(* IEC 61131-3 sources: plc-iiot-stack/src/GVLs/Generated, 1 file *)

(* ---- GVL_IiotMap.gvl.st ---- *)
// AUTO-GENERATED by gen_plc_iiot.py — не редактировать; источник: schema/ (метрики, команды, тревоги)
// Назначение: размеры и таблицы настроек ПЛК-части IIoT-стека КНС-1: метрики телеметрии (топик
//             <site>/<area>/<unit>/<sPath>), белый список команд, тревоги перечня флагмана.
//             Индексы PT_<DEVICE>_<METRIC> — номера метрик в таблице POINT_CFG.
// Документ:   docs/plc_mqtt.md, раздел «Таблицы из схемы данных»
{attribute 'qualified_only'}
VAR_GLOBAL CONSTANT
    POINT_COUNT : DINT := 139;
    RULE_COUNT : DINT := 86;
    CMD_DEVICE_COUNT : DINT := 31;
    ALARM_COUNT : DINT := 88;
    ALARM_WORDS_COUNT : DINT := 28;

    // Метрики (schema/telemetry_catalog.csv)
    PT_P101_RUNNING : DINT := 1;
    PT_P101_STATE : DINT := 2;
    PT_P101_SPEED : DINT := 3;
    PT_P101_SPEED_REF : DINT := 4;
    PT_P101_RUN_HOURS : DINT := 5;
    PT_P101_STARTS : DINT := 6;
    PT_P101_STARTS_LAST_HOUR : DINT := 7;
    PT_P101_RUN_HOURS_MAINT : DINT := 8;
    PT_P101_STARTS_MAINT : DINT := 9;
    PT_P101_VFD_FAULT_CODE : DINT := 10;
    PT_P101_MODE : DINT := 11;
    PT_P101_NE107 : DINT := 12;
    PT_P102_RUNNING : DINT := 13;
    PT_P102_STATE : DINT := 14;
    PT_P102_SPEED : DINT := 15;
    PT_P102_SPEED_REF : DINT := 16;
    PT_P102_RUN_HOURS : DINT := 17;
    PT_P102_STARTS : DINT := 18;
    PT_P102_STARTS_LAST_HOUR : DINT := 19;
    PT_P102_RUN_HOURS_MAINT : DINT := 20;
    PT_P102_STARTS_MAINT : DINT := 21;
    PT_P102_VFD_FAULT_CODE : DINT := 22;
    PT_P102_MODE : DINT := 23;
    PT_P102_NE107 : DINT := 24;
    PT_P103_RUNNING : DINT := 25;
    PT_P103_STATE : DINT := 26;
    PT_P103_SPEED : DINT := 27;
    PT_P103_SPEED_REF : DINT := 28;
    PT_P103_RUN_HOURS : DINT := 29;
    PT_P103_STARTS : DINT := 30;
    PT_P103_STARTS_LAST_HOUR : DINT := 31;
    PT_P103_RUN_HOURS_MAINT : DINT := 32;
    PT_P103_STARTS_MAINT : DINT := 33;
    PT_P103_VFD_FAULT_CODE : DINT := 34;
    PT_P103_MODE : DINT := 35;
    PT_P103_NE107 : DINT := 36;
    PT_V1_RUNNING : DINT := 37;
    PT_V1_STATE : DINT := 38;
    PT_V1_RUN_HOURS : DINT := 39;
    PT_V1_STARTS : DINT := 40;
    PT_V1_STARTS_LAST_HOUR : DINT := 41;
    PT_V1_RUN_HOURS_MAINT : DINT := 42;
    PT_V1_STARTS_MAINT : DINT := 43;
    PT_V1_MODE : DINT := 44;
    PT_V1_NE107 : DINT := 45;
    PT_LT101_LEVEL : DINT := 46;
    PT_LT101_MODE : DINT := 47;
    PT_LT101_NE107 : DINT := 48;
    PT_LS102_LEVEL_HIGH : DINT := 49;
    PT_LS102_MODE : DINT := 50;
    PT_LS102_NE107 : DINT := 51;
    PT_LS103_DRY_RUN : DINT := 52;
    PT_LS103_MODE : DINT := 53;
    PT_LS103_NE107 : DINT := 54;
    PT_IT111_CURRENT : DINT := 55;
    PT_IT111_MODE : DINT := 56;
    PT_IT111_NE107 : DINT := 57;
    PT_TS112_OVERHEAT : DINT := 58;
    PT_TS112_MODE : DINT := 59;
    PT_TS112_NE107 : DINT := 60;
    PT_MS113_LEAK : DINT := 61;
    PT_MS113_MODE : DINT := 62;
    PT_MS113_NE107 : DINT := 63;
    PT_IT121_CURRENT : DINT := 64;
    PT_IT121_MODE : DINT := 65;
    PT_IT121_NE107 : DINT := 66;
    PT_TS122_OVERHEAT : DINT := 67;
    PT_TS122_MODE : DINT := 68;
    PT_TS122_NE107 : DINT := 69;
    PT_MS123_LEAK : DINT := 70;
    PT_MS123_MODE : DINT := 71;
    PT_MS123_NE107 : DINT := 72;
    PT_IT131_CURRENT : DINT := 73;
    PT_IT131_MODE : DINT := 74;
    PT_IT131_NE107 : DINT := 75;
    PT_TS132_OVERHEAT : DINT := 76;
    PT_TS132_MODE : DINT := 77;
    PT_TS132_NE107 : DINT := 78;
    PT_MS133_LEAK : DINT := 79;
    PT_MS133_MODE : DINT := 80;
    PT_MS133_NE107 : DINT := 81;
    PT_PT201_PRESSURE : DINT := 82;
    PT_PT201_MODE : DINT := 83;
    PT_PT201_NE107 : DINT := 84;
    PT_FT202_FLOW : DINT := 85;
    PT_FT202_MODE : DINT := 86;
    PT_FT202_NE107 : DINT := 87;
    PT_LS203_FLOOD : DINT := 88;
    PT_LS203_MODE : DINT := 89;
    PT_LS203_NE107 : DINT := 90;
    PT_ES301_POWER_OK : DINT := 91;
    PT_ES301_MODE : DINT := 92;
    PT_ES301_NE107 : DINT := 93;
    PT_YS302_ON_BATTERY : DINT := 94;
    PT_YS302_MODE : DINT := 95;
    PT_YS302_NE107 : DINT := 96;
    PT_YS303_UPS_FAULT : DINT := 97;
    PT_YS303_MODE : DINT := 98;
    PT_YS303_NE107 : DINT := 99;
    PT_AT401_H2S : DINT := 100;
    PT_AT401_MODE : DINT := 101;
    PT_AT401_NE107 : DINT := 102;
    PT_AT402_CH4 : DINT := 103;
    PT_AT402_MODE : DINT := 104;
    PT_AT402_NE107 : DINT := 105;
    PT_TT403_TEMPERATURE : DINT := 106;
    PT_TT403_MODE : DINT := 107;
    PT_TT403_NE107 : DINT := 108;
    PT_ZS404_DOOR_OPEN : DINT := 109;
    PT_ZS404_MODE : DINT := 110;
    PT_ZS404_NE107 : DINT := 111;
    PT_YS405_FIRE : DINT := 112;
    PT_YS405_MODE : DINT := 113;
    PT_YS405_NE107 : DINT := 114;
    PT_K1_GENERAL_ALARM : DINT := 115;
    PT_KNS1_MODE : DINT := 116;
    PT_KNS1_METHOD : DINT := 117;
    PT_KNS1_CONTROL : DINT := 118;
    PT_KNS1_NE107 : DINT := 119;
    PT_KNS1_STATE : DINT := 120;
    PT_KNS1_PUMPS_REQUIRED : DINT := 121;
    PT_KNS1_PUMPS_RUNNING : DINT := 122;
    PT_KNS1_PUMPS_AVAILABLE : DINT := 123;
    PT_KNS1_LEAD : DINT := 124;
    PT_KNS1_SEQ_REMAIN : DINT := 125;
    PT_KNS1_LEVEL : DINT := 126;
    PT_KNS1_LEVEL_SP : DINT := 127;
    PT_KNS1_SPEED_SP : DINT := 128;
    PT_LIC101_PV : DINT := 129;
    PT_LIC101_SP : DINT := 130;
    PT_LIC101_OUT : DINT := 131;
    PT_LIC101_MODE : DINT := 132;
    PT_LIC101_NE107 : DINT := 133;
    PT_PLC1_UPTIME : DINT := 134;
    PT_PLC1_RECONNECTS : DINT := 135;
    PT_PLC1_QUEUE : DINT := 136;
    PT_PLC1_DROPPED : DINT := 137;
    PT_PLC1_CMD_ACCEPTED : DINT := 138;
    PT_PLC1_CMD_REJECTED : DINT := 139;

    POINT_CFG : ARRAY[1..POINT_COUNT] OF ST_IiotPointCfg := [
        (sPath := 'P101/running', eKind := E_IiotValueKind.Integer, uiDecimals := 0),
        (sPath := 'P101/state', eKind := E_IiotValueKind.Integer, uiDecimals := 0),
        (sPath := 'P101/speed', sUnit := '%', eKind := E_IiotValueKind.Analog, rDeadband := 0.5, uiDecimals := 3),
        (sPath := 'P101/speed_ref', sUnit := '%', eKind := E_IiotValueKind.Analog, rDeadband := 0.5, uiDecimals := 3),
        (sPath := 'P101/run_hours', sUnit := 'h', eKind := E_IiotValueKind.Analog, rDeadband := 0.01, uiDecimals := 3),
        (sPath := 'P101/starts', eKind := E_IiotValueKind.Integer, uiDecimals := 0),
        (sPath := 'P101/starts_last_hour', eKind := E_IiotValueKind.Integer, uiDecimals := 0),
        (sPath := 'P101/run_hours_maint', sUnit := 'h', eKind := E_IiotValueKind.Analog, rDeadband := 0.01,
         uiDecimals := 3),
        (sPath := 'P101/starts_maint', eKind := E_IiotValueKind.Integer, uiDecimals := 0),
        (sPath := 'P101/vfd_fault_code', eKind := E_IiotValueKind.Integer, uiDecimals := 0),
        (sPath := 'P101/mode', eKind := E_IiotValueKind.Integer, uiDecimals := 0),
        (sPath := 'P101/ne107', eKind := E_IiotValueKind.Integer, uiDecimals := 0),
        (sPath := 'P102/running', eKind := E_IiotValueKind.Integer, uiDecimals := 0),
        (sPath := 'P102/state', eKind := E_IiotValueKind.Integer, uiDecimals := 0),
        (sPath := 'P102/speed', sUnit := '%', eKind := E_IiotValueKind.Analog, rDeadband := 0.5, uiDecimals := 3),
        (sPath := 'P102/speed_ref', sUnit := '%', eKind := E_IiotValueKind.Analog, rDeadband := 0.5, uiDecimals := 3),
        (sPath := 'P102/run_hours', sUnit := 'h', eKind := E_IiotValueKind.Analog, rDeadband := 0.01, uiDecimals := 3),
        (sPath := 'P102/starts', eKind := E_IiotValueKind.Integer, uiDecimals := 0),
        (sPath := 'P102/starts_last_hour', eKind := E_IiotValueKind.Integer, uiDecimals := 0),
        (sPath := 'P102/run_hours_maint', sUnit := 'h', eKind := E_IiotValueKind.Analog, rDeadband := 0.01,
         uiDecimals := 3),
        (sPath := 'P102/starts_maint', eKind := E_IiotValueKind.Integer, uiDecimals := 0),
        (sPath := 'P102/vfd_fault_code', eKind := E_IiotValueKind.Integer, uiDecimals := 0),
        (sPath := 'P102/mode', eKind := E_IiotValueKind.Integer, uiDecimals := 0),
        (sPath := 'P102/ne107', eKind := E_IiotValueKind.Integer, uiDecimals := 0),
        (sPath := 'P103/running', eKind := E_IiotValueKind.Integer, uiDecimals := 0),
        (sPath := 'P103/state', eKind := E_IiotValueKind.Integer, uiDecimals := 0),
        (sPath := 'P103/speed', sUnit := '%', eKind := E_IiotValueKind.Analog, rDeadband := 0.5, uiDecimals := 3),
        (sPath := 'P103/speed_ref', sUnit := '%', eKind := E_IiotValueKind.Analog, rDeadband := 0.5, uiDecimals := 3),
        (sPath := 'P103/run_hours', sUnit := 'h', eKind := E_IiotValueKind.Analog, rDeadband := 0.01, uiDecimals := 3),
        (sPath := 'P103/starts', eKind := E_IiotValueKind.Integer, uiDecimals := 0),
        (sPath := 'P103/starts_last_hour', eKind := E_IiotValueKind.Integer, uiDecimals := 0),
        (sPath := 'P103/run_hours_maint', sUnit := 'h', eKind := E_IiotValueKind.Analog, rDeadband := 0.01,
         uiDecimals := 3),
        (sPath := 'P103/starts_maint', eKind := E_IiotValueKind.Integer, uiDecimals := 0),
        (sPath := 'P103/vfd_fault_code', eKind := E_IiotValueKind.Integer, uiDecimals := 0),
        (sPath := 'P103/mode', eKind := E_IiotValueKind.Integer, uiDecimals := 0),
        (sPath := 'P103/ne107', eKind := E_IiotValueKind.Integer, uiDecimals := 0),
        (sPath := 'V1/running', eKind := E_IiotValueKind.Integer, uiDecimals := 0),
        (sPath := 'V1/state', eKind := E_IiotValueKind.Integer, uiDecimals := 0),
        (sPath := 'V1/run_hours', sUnit := 'h', eKind := E_IiotValueKind.Analog, rDeadband := 0.01, uiDecimals := 3),
        (sPath := 'V1/starts', eKind := E_IiotValueKind.Integer, uiDecimals := 0),
        (sPath := 'V1/starts_last_hour', eKind := E_IiotValueKind.Integer, uiDecimals := 0),
        (sPath := 'V1/run_hours_maint', sUnit := 'h', eKind := E_IiotValueKind.Analog, rDeadband := 0.01,
         uiDecimals := 3),
        (sPath := 'V1/starts_maint', eKind := E_IiotValueKind.Integer, uiDecimals := 0),
        (sPath := 'V1/mode', eKind := E_IiotValueKind.Integer, uiDecimals := 0),
        (sPath := 'V1/ne107', eKind := E_IiotValueKind.Integer, uiDecimals := 0),
        (sPath := 'LT101/level', sUnit := 'm', eKind := E_IiotValueKind.Analog, rDeadband := 0.01, uiDecimals := 3),
        (sPath := 'LT101/mode', eKind := E_IiotValueKind.Integer, uiDecimals := 0),
        (sPath := 'LT101/ne107', eKind := E_IiotValueKind.Integer, uiDecimals := 0),
        (sPath := 'LS102/level_high', eKind := E_IiotValueKind.Integer, uiDecimals := 0),
        (sPath := 'LS102/mode', eKind := E_IiotValueKind.Integer, uiDecimals := 0),
        (sPath := 'LS102/ne107', eKind := E_IiotValueKind.Integer, uiDecimals := 0),
        (sPath := 'LS103/dry_run', eKind := E_IiotValueKind.Integer, uiDecimals := 0),
        (sPath := 'LS103/mode', eKind := E_IiotValueKind.Integer, uiDecimals := 0),
        (sPath := 'LS103/ne107', eKind := E_IiotValueKind.Integer, uiDecimals := 0),
        (sPath := 'IT111/current', sUnit := 'A', eKind := E_IiotValueKind.Analog, rDeadband := 0.2, uiDecimals := 3),
        (sPath := 'IT111/mode', eKind := E_IiotValueKind.Integer, uiDecimals := 0),
        (sPath := 'IT111/ne107', eKind := E_IiotValueKind.Integer, uiDecimals := 0),
        (sPath := 'TS112/overheat', eKind := E_IiotValueKind.Integer, uiDecimals := 0),
        (sPath := 'TS112/mode', eKind := E_IiotValueKind.Integer, uiDecimals := 0),
        (sPath := 'TS112/ne107', eKind := E_IiotValueKind.Integer, uiDecimals := 0),
        (sPath := 'MS113/leak', eKind := E_IiotValueKind.Integer, uiDecimals := 0),
        (sPath := 'MS113/mode', eKind := E_IiotValueKind.Integer, uiDecimals := 0),
        (sPath := 'MS113/ne107', eKind := E_IiotValueKind.Integer, uiDecimals := 0),
        (sPath := 'IT121/current', sUnit := 'A', eKind := E_IiotValueKind.Analog, rDeadband := 0.2, uiDecimals := 3),
        (sPath := 'IT121/mode', eKind := E_IiotValueKind.Integer, uiDecimals := 0),
        (sPath := 'IT121/ne107', eKind := E_IiotValueKind.Integer, uiDecimals := 0),
        (sPath := 'TS122/overheat', eKind := E_IiotValueKind.Integer, uiDecimals := 0),
        (sPath := 'TS122/mode', eKind := E_IiotValueKind.Integer, uiDecimals := 0),
        (sPath := 'TS122/ne107', eKind := E_IiotValueKind.Integer, uiDecimals := 0),
        (sPath := 'MS123/leak', eKind := E_IiotValueKind.Integer, uiDecimals := 0),
        (sPath := 'MS123/mode', eKind := E_IiotValueKind.Integer, uiDecimals := 0),
        (sPath := 'MS123/ne107', eKind := E_IiotValueKind.Integer, uiDecimals := 0),
        (sPath := 'IT131/current', sUnit := 'A', eKind := E_IiotValueKind.Analog, rDeadband := 0.2, uiDecimals := 3),
        (sPath := 'IT131/mode', eKind := E_IiotValueKind.Integer, uiDecimals := 0),
        (sPath := 'IT131/ne107', eKind := E_IiotValueKind.Integer, uiDecimals := 0),
        (sPath := 'TS132/overheat', eKind := E_IiotValueKind.Integer, uiDecimals := 0),
        (sPath := 'TS132/mode', eKind := E_IiotValueKind.Integer, uiDecimals := 0),
        (sPath := 'TS132/ne107', eKind := E_IiotValueKind.Integer, uiDecimals := 0),
        (sPath := 'MS133/leak', eKind := E_IiotValueKind.Integer, uiDecimals := 0),
        (sPath := 'MS133/mode', eKind := E_IiotValueKind.Integer, uiDecimals := 0),
        (sPath := 'MS133/ne107', eKind := E_IiotValueKind.Integer, uiDecimals := 0),
        (sPath := 'PT201/pressure', sUnit := 'bar', eKind := E_IiotValueKind.Analog, rDeadband := 0.02,
         uiDecimals := 3),
        (sPath := 'PT201/mode', eKind := E_IiotValueKind.Integer, uiDecimals := 0),
        (sPath := 'PT201/ne107', eKind := E_IiotValueKind.Integer, uiDecimals := 0),
        (sPath := 'FT202/flow', sUnit := 'm3/h', eKind := E_IiotValueKind.Analog, rDeadband := 2.0, uiDecimals := 3),
        (sPath := 'FT202/mode', eKind := E_IiotValueKind.Integer, uiDecimals := 0),
        (sPath := 'FT202/ne107', eKind := E_IiotValueKind.Integer, uiDecimals := 0),
        (sPath := 'LS203/flood', eKind := E_IiotValueKind.Integer, uiDecimals := 0),
        (sPath := 'LS203/mode', eKind := E_IiotValueKind.Integer, uiDecimals := 0),
        (sPath := 'LS203/ne107', eKind := E_IiotValueKind.Integer, uiDecimals := 0),
        (sPath := 'ES301/power_ok', eKind := E_IiotValueKind.Integer, uiDecimals := 0),
        (sPath := 'ES301/mode', eKind := E_IiotValueKind.Integer, uiDecimals := 0),
        (sPath := 'ES301/ne107', eKind := E_IiotValueKind.Integer, uiDecimals := 0),
        (sPath := 'YS302/on_battery', eKind := E_IiotValueKind.Integer, uiDecimals := 0),
        (sPath := 'YS302/mode', eKind := E_IiotValueKind.Integer, uiDecimals := 0),
        (sPath := 'YS302/ne107', eKind := E_IiotValueKind.Integer, uiDecimals := 0),
        (sPath := 'YS303/ups_fault', eKind := E_IiotValueKind.Integer, uiDecimals := 0),
        (sPath := 'YS303/mode', eKind := E_IiotValueKind.Integer, uiDecimals := 0),
        (sPath := 'YS303/ne107', eKind := E_IiotValueKind.Integer, uiDecimals := 0),
        (sPath := 'AT401/h2s', sUnit := 'mg/m3', eKind := E_IiotValueKind.Analog, rDeadband := 0.2, uiDecimals := 3),
        (sPath := 'AT401/mode', eKind := E_IiotValueKind.Integer, uiDecimals := 0),
        (sPath := 'AT401/ne107', eKind := E_IiotValueKind.Integer, uiDecimals := 0),
        (sPath := 'AT402/ch4', sUnit := '%LEL', eKind := E_IiotValueKind.Analog, rDeadband := 0.5, uiDecimals := 3),
        (sPath := 'AT402/mode', eKind := E_IiotValueKind.Integer, uiDecimals := 0),
        (sPath := 'AT402/ne107', eKind := E_IiotValueKind.Integer, uiDecimals := 0),
        (sPath := 'TT403/temperature', sUnit := 'degC', eKind := E_IiotValueKind.Analog, rDeadband := 0.2,
         uiDecimals := 3),
        (sPath := 'TT403/mode', eKind := E_IiotValueKind.Integer, uiDecimals := 0),
        (sPath := 'TT403/ne107', eKind := E_IiotValueKind.Integer, uiDecimals := 0),
        (sPath := 'ZS404/door_open', eKind := E_IiotValueKind.Integer, uiDecimals := 0),
        (sPath := 'ZS404/mode', eKind := E_IiotValueKind.Integer, uiDecimals := 0),
        (sPath := 'ZS404/ne107', eKind := E_IiotValueKind.Integer, uiDecimals := 0),
        (sPath := 'YS405/fire', eKind := E_IiotValueKind.Integer, uiDecimals := 0),
        (sPath := 'YS405/mode', eKind := E_IiotValueKind.Integer, uiDecimals := 0),
        (sPath := 'YS405/ne107', eKind := E_IiotValueKind.Integer, uiDecimals := 0),
        (sPath := 'K1/general_alarm', eKind := E_IiotValueKind.Integer, uiDecimals := 0),
        (sPath := 'KNS1/mode', eKind := E_IiotValueKind.Integer, uiDecimals := 0),
        (sPath := 'KNS1/method', eKind := E_IiotValueKind.Integer, uiDecimals := 0),
        (sPath := 'KNS1/control', eKind := E_IiotValueKind.Integer, uiDecimals := 0),
        (sPath := 'KNS1/ne107', eKind := E_IiotValueKind.Integer, uiDecimals := 0),
        (sPath := 'KNS1/state', eKind := E_IiotValueKind.Integer, uiDecimals := 0),
        (sPath := 'KNS1/pumps_required', eKind := E_IiotValueKind.Integer, uiDecimals := 0),
        (sPath := 'KNS1/pumps_running', eKind := E_IiotValueKind.Integer, uiDecimals := 0),
        (sPath := 'KNS1/pumps_available', eKind := E_IiotValueKind.Integer, uiDecimals := 0),
        (sPath := 'KNS1/lead', eKind := E_IiotValueKind.Integer, uiDecimals := 0),
        (sPath := 'KNS1/seq_remain', sUnit := 's', eKind := E_IiotValueKind.Integer, uiDecimals := 0),
        (sPath := 'KNS1/level', sUnit := 'm', eKind := E_IiotValueKind.Analog, rDeadband := 0.01, uiDecimals := 3),
        (sPath := 'KNS1/level_sp', sUnit := 'm', eKind := E_IiotValueKind.Analog, rDeadband := 0.01, uiDecimals := 3),
        (sPath := 'KNS1/speed_sp', sUnit := '%', eKind := E_IiotValueKind.Analog, rDeadband := 0.5, uiDecimals := 3),
        (sPath := 'LIC101/pv', sUnit := 'm', eKind := E_IiotValueKind.Analog, rDeadband := 0.01, uiDecimals := 3),
        (sPath := 'LIC101/sp', sUnit := 'm', eKind := E_IiotValueKind.Analog, rDeadband := 0.01, uiDecimals := 3),
        (sPath := 'LIC101/out', sUnit := '%', eKind := E_IiotValueKind.Analog, rDeadband := 0.5, uiDecimals := 3),
        (sPath := 'LIC101/mode', eKind := E_IiotValueKind.Integer, uiDecimals := 0),
        (sPath := 'LIC101/ne107', eKind := E_IiotValueKind.Integer, uiDecimals := 0),
        (sPath := 'PLC1/uptime', sUnit := 's', eKind := E_IiotValueKind.Integer, uiDecimals := 0,
         xPeriodicOnly := TRUE),
        (sPath := 'PLC1/reconnects', eKind := E_IiotValueKind.Integer, uiDecimals := 0),
        (sPath := 'PLC1/queue', eKind := E_IiotValueKind.Integer, uiDecimals := 0),
        (sPath := 'PLC1/dropped', eKind := E_IiotValueKind.Integer, uiDecimals := 0),
        (sPath := 'PLC1/cmd_accepted', eKind := E_IiotValueKind.Integer, uiDecimals := 0),
        (sPath := 'PLC1/cmd_rejected', eKind := E_IiotValueKind.Integer, uiDecimals := 0)];

    // Белый список команд (schema/command_whitelist.csv)
    RULE_CFG : ARRAY[1..RULE_COUNT] OF ST_IiotCmdRule := [
        (sDevice := 'P101', eCommand := E_IiotCommand.SetAuto, diDev := 1),
        (sDevice := 'P101', eCommand := E_IiotCommand.SetManual, diDev := 1),
        (sDevice := 'P101', eCommand := E_IiotCommand.Start, diDev := 1),
        (sDevice := 'P101', eCommand := E_IiotCommand.Stop, diDev := 1),
        (sDevice := 'P101', eCommand := E_IiotCommand.SpeedSp, xRange := TRUE, rMin := 0.0, rMax := 100.0, diDev := 1),
        (sDevice := 'P101', eCommand := E_IiotCommand.Ack, diDev := 1),
        (sDevice := 'P101', eCommand := E_IiotCommand.Reset, diDev := 1),
        (sDevice := 'P102', eCommand := E_IiotCommand.SetAuto, diDev := 2),
        (sDevice := 'P102', eCommand := E_IiotCommand.SetManual, diDev := 2),
        (sDevice := 'P102', eCommand := E_IiotCommand.Start, diDev := 2),
        (sDevice := 'P102', eCommand := E_IiotCommand.Stop, diDev := 2),
        (sDevice := 'P102', eCommand := E_IiotCommand.SpeedSp, xRange := TRUE, rMin := 0.0, rMax := 100.0, diDev := 2),
        (sDevice := 'P102', eCommand := E_IiotCommand.Ack, diDev := 2),
        (sDevice := 'P102', eCommand := E_IiotCommand.Reset, diDev := 2),
        (sDevice := 'P103', eCommand := E_IiotCommand.SetAuto, diDev := 3),
        (sDevice := 'P103', eCommand := E_IiotCommand.SetManual, diDev := 3),
        (sDevice := 'P103', eCommand := E_IiotCommand.Start, diDev := 3),
        (sDevice := 'P103', eCommand := E_IiotCommand.Stop, diDev := 3),
        (sDevice := 'P103', eCommand := E_IiotCommand.SpeedSp, xRange := TRUE, rMin := 0.0, rMax := 100.0, diDev := 3),
        (sDevice := 'P103', eCommand := E_IiotCommand.Ack, diDev := 3),
        (sDevice := 'P103', eCommand := E_IiotCommand.Reset, diDev := 3),
        (sDevice := 'V1', eCommand := E_IiotCommand.SetAuto, diDev := 4),
        (sDevice := 'V1', eCommand := E_IiotCommand.SetManual, diDev := 4),
        (sDevice := 'V1', eCommand := E_IiotCommand.Start, diDev := 4),
        (sDevice := 'V1', eCommand := E_IiotCommand.Stop, diDev := 4),
        (sDevice := 'V1', eCommand := E_IiotCommand.Ack, diDev := 4),
        (sDevice := 'V1', eCommand := E_IiotCommand.Reset, diDev := 4),
        (sDevice := 'LT101', eCommand := E_IiotCommand.Ack, diDev := 5),
        (sDevice := 'LT101', eCommand := E_IiotCommand.Reset, diDev := 5),
        (sDevice := 'LS102', eCommand := E_IiotCommand.Ack, diDev := 6),
        (sDevice := 'LS102', eCommand := E_IiotCommand.Reset, diDev := 6),
        (sDevice := 'LS103', eCommand := E_IiotCommand.Ack, diDev := 7),
        (sDevice := 'LS103', eCommand := E_IiotCommand.Reset, diDev := 7),
        (sDevice := 'IT111', eCommand := E_IiotCommand.Ack, diDev := 8),
        (sDevice := 'IT111', eCommand := E_IiotCommand.Reset, diDev := 8),
        (sDevice := 'TS112', eCommand := E_IiotCommand.Ack, diDev := 9),
        (sDevice := 'TS112', eCommand := E_IiotCommand.Reset, diDev := 9),
        (sDevice := 'MS113', eCommand := E_IiotCommand.Ack, diDev := 10),
        (sDevice := 'MS113', eCommand := E_IiotCommand.Reset, diDev := 10),
        (sDevice := 'IT121', eCommand := E_IiotCommand.Ack, diDev := 11),
        (sDevice := 'IT121', eCommand := E_IiotCommand.Reset, diDev := 11),
        (sDevice := 'TS122', eCommand := E_IiotCommand.Ack, diDev := 12),
        (sDevice := 'TS122', eCommand := E_IiotCommand.Reset, diDev := 12),
        (sDevice := 'MS123', eCommand := E_IiotCommand.Ack, diDev := 13),
        (sDevice := 'MS123', eCommand := E_IiotCommand.Reset, diDev := 13),
        (sDevice := 'IT131', eCommand := E_IiotCommand.Ack, diDev := 14),
        (sDevice := 'IT131', eCommand := E_IiotCommand.Reset, diDev := 14),
        (sDevice := 'TS132', eCommand := E_IiotCommand.Ack, diDev := 15),
        (sDevice := 'TS132', eCommand := E_IiotCommand.Reset, diDev := 15),
        (sDevice := 'MS133', eCommand := E_IiotCommand.Ack, diDev := 16),
        (sDevice := 'MS133', eCommand := E_IiotCommand.Reset, diDev := 16),
        (sDevice := 'PT201', eCommand := E_IiotCommand.Ack, diDev := 17),
        (sDevice := 'PT201', eCommand := E_IiotCommand.Reset, diDev := 17),
        (sDevice := 'FT202', eCommand := E_IiotCommand.Ack, diDev := 18),
        (sDevice := 'FT202', eCommand := E_IiotCommand.Reset, diDev := 18),
        (sDevice := 'LS203', eCommand := E_IiotCommand.Ack, diDev := 19),
        (sDevice := 'LS203', eCommand := E_IiotCommand.Reset, diDev := 19),
        (sDevice := 'ES301', eCommand := E_IiotCommand.Ack, diDev := 20),
        (sDevice := 'ES301', eCommand := E_IiotCommand.Reset, diDev := 20),
        (sDevice := 'YS302', eCommand := E_IiotCommand.Ack, diDev := 21),
        (sDevice := 'YS302', eCommand := E_IiotCommand.Reset, diDev := 21),
        (sDevice := 'YS303', eCommand := E_IiotCommand.Ack, diDev := 22),
        (sDevice := 'YS303', eCommand := E_IiotCommand.Reset, diDev := 22),
        (sDevice := 'AT401', eCommand := E_IiotCommand.Ack, diDev := 23),
        (sDevice := 'AT401', eCommand := E_IiotCommand.Reset, diDev := 23),
        (sDevice := 'AT402', eCommand := E_IiotCommand.Ack, diDev := 24),
        (sDevice := 'AT402', eCommand := E_IiotCommand.Reset, diDev := 24),
        (sDevice := 'TT403', eCommand := E_IiotCommand.Ack, diDev := 25),
        (sDevice := 'TT403', eCommand := E_IiotCommand.Reset, diDev := 25),
        (sDevice := 'ZS404', eCommand := E_IiotCommand.Ack, diDev := 26),
        (sDevice := 'ZS404', eCommand := E_IiotCommand.Reset, diDev := 26),
        (sDevice := 'YS405', eCommand := E_IiotCommand.Ack, diDev := 27),
        (sDevice := 'YS405', eCommand := E_IiotCommand.Reset, diDev := 27),
        (sDevice := 'HS501', eCommand := E_IiotCommand.Ack, diDev := 28),
        (sDevice := 'HS501', eCommand := E_IiotCommand.Reset, diDev := 28),
        (sDevice := 'HS502', eCommand := E_IiotCommand.Ack, diDev := 29),
        (sDevice := 'HS502', eCommand := E_IiotCommand.Reset, diDev := 29),
        (sDevice := 'KNS1', eCommand := E_IiotCommand.SetAuto, diDev := 30),
        (sDevice := 'KNS1', eCommand := E_IiotCommand.SetManual, diDev := 30),
        (sDevice := 'KNS1', eCommand := E_IiotCommand.SetStepped, diDev := 30),
        (sDevice := 'KNS1', eCommand := E_IiotCommand.SetLevelPid, diDev := 30),
        (sDevice := 'KNS1', eCommand := E_IiotCommand.AckAll, diDev := 30),
        (sDevice := 'KNS1', eCommand := E_IiotCommand.ResetAll, diDev := 30),
        (sDevice := 'KNS1', eCommand := E_IiotCommand.Silence, diDev := 30),
        (sDevice := 'LIC101', eCommand := E_IiotCommand.SetAuto, diDev := 31),
        (sDevice := 'LIC101', eCommand := E_IiotCommand.SetManual, diDev := 31)];

    // Тревоги (schema/source/scada_alarms.csv, station_alarms.csv): uiSlot — бит в словах тревог,
    // diWords — строка таблицы слов устройства
    ALARM_CFG : ARRAY[1..ALARM_COUNT] OF ST_IiotAlarmCfg := [
        (udiId := 110, sDevice := 'P101', sSuffix := 'FTS', uiSlot := 0, ePriority := E_IiotAlarmPriority.Medium,
         diWords := 1),
        (udiId := 111, sDevice := 'P101', sSuffix := 'FBL', uiSlot := 1, ePriority := E_IiotAlarmPriority.Medium,
         diWords := 1),
        (udiId := 112, sDevice := 'P101', sSuffix := 'FTP', uiSlot := 2, ePriority := E_IiotAlarmPriority.High,
         diWords := 1),
        (udiId := 113, sDevice := 'P101', sSuffix := 'UCR', uiSlot := 3, ePriority := E_IiotAlarmPriority.High,
         diWords := 1),
        (udiId := 114, sDevice := 'P101', sSuffix := 'EXT', uiSlot := 4, ePriority := E_IiotAlarmPriority.Medium,
         diWords := 1),
        (udiId := 116, sDevice := 'P101', sSuffix := 'COM', uiSlot := 6, ePriority := E_IiotAlarmPriority.Medium,
         diWords := 1),
        (udiId := 117, sDevice := 'P101', sSuffix := 'SPD', uiSlot := 7, ePriority := E_IiotAlarmPriority.Low,
         diWords := 1),
        (udiId := 120, sDevice := 'P102', sSuffix := 'FTS', uiSlot := 0, ePriority := E_IiotAlarmPriority.Medium,
         diWords := 2),
        (udiId := 121, sDevice := 'P102', sSuffix := 'FBL', uiSlot := 1, ePriority := E_IiotAlarmPriority.Medium,
         diWords := 2),
        (udiId := 122, sDevice := 'P102', sSuffix := 'FTP', uiSlot := 2, ePriority := E_IiotAlarmPriority.High,
         diWords := 2),
        (udiId := 123, sDevice := 'P102', sSuffix := 'UCR', uiSlot := 3, ePriority := E_IiotAlarmPriority.High,
         diWords := 2),
        (udiId := 124, sDevice := 'P102', sSuffix := 'EXT', uiSlot := 4, ePriority := E_IiotAlarmPriority.Medium,
         diWords := 2),
        (udiId := 126, sDevice := 'P102', sSuffix := 'COM', uiSlot := 6, ePriority := E_IiotAlarmPriority.Medium,
         diWords := 2),
        (udiId := 127, sDevice := 'P102', sSuffix := 'SPD', uiSlot := 7, ePriority := E_IiotAlarmPriority.Low,
         diWords := 2),
        (udiId := 130, sDevice := 'P103', sSuffix := 'FTS', uiSlot := 0, ePriority := E_IiotAlarmPriority.Medium,
         diWords := 3),
        (udiId := 131, sDevice := 'P103', sSuffix := 'FBL', uiSlot := 1, ePriority := E_IiotAlarmPriority.Medium,
         diWords := 3),
        (udiId := 132, sDevice := 'P103', sSuffix := 'FTP', uiSlot := 2, ePriority := E_IiotAlarmPriority.High,
         diWords := 3),
        (udiId := 133, sDevice := 'P103', sSuffix := 'UCR', uiSlot := 3, ePriority := E_IiotAlarmPriority.High,
         diWords := 3),
        (udiId := 134, sDevice := 'P103', sSuffix := 'EXT', uiSlot := 4, ePriority := E_IiotAlarmPriority.Medium,
         diWords := 3),
        (udiId := 136, sDevice := 'P103', sSuffix := 'COM', uiSlot := 6, ePriority := E_IiotAlarmPriority.Medium,
         diWords := 3),
        (udiId := 137, sDevice := 'P103', sSuffix := 'SPD', uiSlot := 7, ePriority := E_IiotAlarmPriority.Low,
         diWords := 3),
        (udiId := 140, sDevice := 'V1', sSuffix := 'FTS', uiSlot := 0, ePriority := E_IiotAlarmPriority.Low,
         diWords := 4),
        (udiId := 141, sDevice := 'V1', sSuffix := 'FBL', uiSlot := 1, ePriority := E_IiotAlarmPriority.Low,
         diWords := 4),
        (udiId := 142, sDevice := 'V1', sSuffix := 'FTP', uiSlot := 2, ePriority := E_IiotAlarmPriority.High,
         diWords := 4),
        (udiId := 143, sDevice := 'V1', sSuffix := 'UCR', uiSlot := 3, ePriority := E_IiotAlarmPriority.High,
         diWords := 4),
        (udiId := 144, sDevice := 'V1', sSuffix := 'EXT', uiSlot := 4, ePriority := E_IiotAlarmPriority.Low,
         diWords := 4),
        (udiId := 1010, sDevice := 'LT101', sSuffix := 'HH', uiSlot := 0, ePriority := E_IiotAlarmPriority.High,
         diWords := 5),
        (udiId := 1011, sDevice := 'LT101', sSuffix := 'H', uiSlot := 1, ePriority := E_IiotAlarmPriority.Medium,
         diWords := 5),
        (udiId := 1012, sDevice := 'LT101', sSuffix := 'L', uiSlot := 2, ePriority := E_IiotAlarmPriority.Medium,
         diWords := 5),
        (udiId := 1013, sDevice := 'LT101', sSuffix := 'LL', uiSlot := 3, ePriority := E_IiotAlarmPriority.High,
         diWords := 5),
        (udiId := 1014, sDevice := 'LT101', sSuffix := 'FAIL', uiSlot := 4, ePriority := E_IiotAlarmPriority.Medium,
         diWords := 5),
        (udiId := 1015, sDevice := 'LT101', sSuffix := 'OOR', uiSlot := 5, ePriority := E_IiotAlarmPriority.Low,
         diWords := 5),
        (udiId := 1020, sDevice := 'LS102', sSuffix := 'ALM', uiSlot := 0, ePriority := E_IiotAlarmPriority.High,
         diWords := 6),
        (udiId := 1030, sDevice := 'LS103', sSuffix := 'ALM', uiSlot := 0, ePriority := E_IiotAlarmPriority.High,
         diWords := 7),
        (udiId := 1110, sDevice := 'IT111', sSuffix := 'HH', uiSlot := 0, ePriority := E_IiotAlarmPriority.Medium,
         diWords := 8),
        (udiId := 1111, sDevice := 'IT111', sSuffix := 'H', uiSlot := 1, ePriority := E_IiotAlarmPriority.Low,
         diWords := 8),
        (udiId := 1114, sDevice := 'IT111', sSuffix := 'FAIL', uiSlot := 4, ePriority := E_IiotAlarmPriority.Medium,
         diWords := 8),
        (udiId := 1120, sDevice := 'TS112', sSuffix := 'ALM', uiSlot := 0, ePriority := E_IiotAlarmPriority.High,
         diWords := 9),
        (udiId := 1130, sDevice := 'MS113', sSuffix := 'ALM', uiSlot := 0, ePriority := E_IiotAlarmPriority.Medium,
         diWords := 10),
        (udiId := 1210, sDevice := 'IT121', sSuffix := 'HH', uiSlot := 0, ePriority := E_IiotAlarmPriority.Medium,
         diWords := 11),
        (udiId := 1211, sDevice := 'IT121', sSuffix := 'H', uiSlot := 1, ePriority := E_IiotAlarmPriority.Low,
         diWords := 11),
        (udiId := 1214, sDevice := 'IT121', sSuffix := 'FAIL', uiSlot := 4, ePriority := E_IiotAlarmPriority.Medium,
         diWords := 11),
        (udiId := 1220, sDevice := 'TS122', sSuffix := 'ALM', uiSlot := 0, ePriority := E_IiotAlarmPriority.High,
         diWords := 12),
        (udiId := 1230, sDevice := 'MS123', sSuffix := 'ALM', uiSlot := 0, ePriority := E_IiotAlarmPriority.Medium,
         diWords := 13),
        (udiId := 1310, sDevice := 'IT131', sSuffix := 'HH', uiSlot := 0, ePriority := E_IiotAlarmPriority.Medium,
         diWords := 14),
        (udiId := 1311, sDevice := 'IT131', sSuffix := 'H', uiSlot := 1, ePriority := E_IiotAlarmPriority.Low,
         diWords := 14),
        (udiId := 1314, sDevice := 'IT131', sSuffix := 'FAIL', uiSlot := 4, ePriority := E_IiotAlarmPriority.Medium,
         diWords := 14),
        (udiId := 1320, sDevice := 'TS132', sSuffix := 'ALM', uiSlot := 0, ePriority := E_IiotAlarmPriority.High,
         diWords := 15),
        (udiId := 1330, sDevice := 'MS133', sSuffix := 'ALM', uiSlot := 0, ePriority := E_IiotAlarmPriority.Medium,
         diWords := 16),
        (udiId := 2010, sDevice := 'PT201', sSuffix := 'HH', uiSlot := 0, ePriority := E_IiotAlarmPriority.High,
         diWords := 17),
        (udiId := 2011, sDevice := 'PT201', sSuffix := 'H', uiSlot := 1, ePriority := E_IiotAlarmPriority.Medium,
         diWords := 17),
        (udiId := 2012, sDevice := 'PT201', sSuffix := 'L', uiSlot := 2, ePriority := E_IiotAlarmPriority.Medium,
         diWords := 17),
        (udiId := 2013, sDevice := 'PT201', sSuffix := 'LL', uiSlot := 3, ePriority := E_IiotAlarmPriority.High,
         diWords := 17),
        (udiId := 2014, sDevice := 'PT201', sSuffix := 'FAIL', uiSlot := 4, ePriority := E_IiotAlarmPriority.Medium,
         diWords := 17),
        (udiId := 2015, sDevice := 'PT201', sSuffix := 'OOR', uiSlot := 5, ePriority := E_IiotAlarmPriority.Low,
         diWords := 17),
        (udiId := 2022, sDevice := 'FT202', sSuffix := 'L', uiSlot := 2, ePriority := E_IiotAlarmPriority.Medium,
         diWords := 18),
        (udiId := 2024, sDevice := 'FT202', sSuffix := 'FAIL', uiSlot := 4, ePriority := E_IiotAlarmPriority.Medium,
         diWords := 18),
        (udiId := 2025, sDevice := 'FT202', sSuffix := 'OOR', uiSlot := 5, ePriority := E_IiotAlarmPriority.Low,
         diWords := 18),
        (udiId := 2030, sDevice := 'LS203', sSuffix := 'ALM', uiSlot := 0, ePriority := E_IiotAlarmPriority.Medium,
         diWords := 19),
        (udiId := 3010, sDevice := 'ES301', sSuffix := 'ALM', uiSlot := 0, ePriority := E_IiotAlarmPriority.High,
         diWords := 20),
        (udiId := 3020, sDevice := 'YS302', sSuffix := 'ALM', uiSlot := 0, ePriority := E_IiotAlarmPriority.Medium,
         diWords := 21),
        (udiId := 3030, sDevice := 'YS303', sSuffix := 'ALM', uiSlot := 0, ePriority := E_IiotAlarmPriority.Medium,
         diWords := 22),
        (udiId := 4010, sDevice := 'AT401', sSuffix := 'HH', uiSlot := 0, ePriority := E_IiotAlarmPriority.High,
         diWords := 23),
        (udiId := 4011, sDevice := 'AT401', sSuffix := 'H', uiSlot := 1, ePriority := E_IiotAlarmPriority.Medium,
         diWords := 23),
        (udiId := 4014, sDevice := 'AT401', sSuffix := 'FAIL', uiSlot := 4, ePriority := E_IiotAlarmPriority.Medium,
         diWords := 23),
        (udiId := 4015, sDevice := 'AT401', sSuffix := 'OOR', uiSlot := 5, ePriority := E_IiotAlarmPriority.Low,
         diWords := 23),
        (udiId := 4020, sDevice := 'AT402', sSuffix := 'HH', uiSlot := 0, ePriority := E_IiotAlarmPriority.High,
         diWords := 24),
        (udiId := 4021, sDevice := 'AT402', sSuffix := 'H', uiSlot := 1, ePriority := E_IiotAlarmPriority.Medium,
         diWords := 24),
        (udiId := 4024, sDevice := 'AT402', sSuffix := 'FAIL', uiSlot := 4, ePriority := E_IiotAlarmPriority.Medium,
         diWords := 24),
        (udiId := 4025, sDevice := 'AT402', sSuffix := 'OOR', uiSlot := 5, ePriority := E_IiotAlarmPriority.Low,
         diWords := 24),
        (udiId := 4031, sDevice := 'TT403', sSuffix := 'H', uiSlot := 1, ePriority := E_IiotAlarmPriority.Low,
         diWords := 25),
        (udiId := 4032, sDevice := 'TT403', sSuffix := 'L', uiSlot := 2, ePriority := E_IiotAlarmPriority.Low,
         diWords := 25),
        (udiId := 4034, sDevice := 'TT403', sSuffix := 'FAIL', uiSlot := 4, ePriority := E_IiotAlarmPriority.Medium,
         diWords := 25),
        (udiId := 4040, sDevice := 'ZS404', sSuffix := 'ALM', uiSlot := 0, ePriority := E_IiotAlarmPriority.Low,
         diWords := 26),
        (udiId := 4050, sDevice := 'YS405', sSuffix := 'ALM', uiSlot := 0, ePriority := E_IiotAlarmPriority.High,
         diWords := 27),
        (udiId := 100001, sDevice := 'KNS1', sSuffix := 'EHL', uiSlot := 0, ePriority := E_IiotAlarmPriority.Critical,
         diWords := 28),
        (udiId := 100002, sDevice := 'KNS1', sSuffix := 'DRY', uiSlot := 1, ePriority := E_IiotAlarmPriority.High,
         diWords := 28),
        (udiId := 100003, sDevice := 'KNS1', sSuffix := 'LACK', uiSlot := 2, ePriority := E_IiotAlarmPriority.High,
         diWords := 28),
        (udiId := 100004, sDevice := 'KNS1', sSuffix := 'NORES', uiSlot := 3, ePriority := E_IiotAlarmPriority.High,
         diWords := 28),
        (udiId := 100005, sDevice := 'KNS1', sSuffix := 'ATS', uiSlot := 4, ePriority := E_IiotAlarmPriority.Medium,
         diWords := 28),
        (udiId := 100006, sDevice := 'KNS1', sSuffix := 'FLOAT', uiSlot := 5, ePriority := E_IiotAlarmPriority.Medium,
         diWords := 28),
        (udiId := 100007, sDevice := 'KNS1', sSuffix := 'LDEV', uiSlot := 6, ePriority := E_IiotAlarmPriority.Medium,
         diWords := 28),
        (udiId := 100008, sDevice := 'KNS1', sSuffix := 'STEP', uiSlot := 7, ePriority := E_IiotAlarmPriority.Low,
         diWords := 28),
        (udiId := 100009, sDevice := 'KNS1', sSuffix := 'NOAUTO', uiSlot := 8, ePriority := E_IiotAlarmPriority.Low,
         diWords := 28),
        (udiId := 100010, sDevice := 'KNS1', sSuffix := 'UL1', uiSlot := 9, ePriority := E_IiotAlarmPriority.Medium,
         diWords := 28),
        (udiId := 100011, sDevice := 'KNS1', sSuffix := 'UL2', uiSlot := 10, ePriority := E_IiotAlarmPriority.Medium,
         diWords := 28),
        (udiId := 100012, sDevice := 'KNS1', sSuffix := 'UL3', uiSlot := 11, ePriority := E_IiotAlarmPriority.Medium,
         diWords := 28),
        (udiId := 100013, sDevice := 'KNS1', sSuffix := 'SIM', uiSlot := 12, ePriority := E_IiotAlarmPriority.Low,
         diWords := 28)];
END_VAR
